(* IEC 61131-3 sources: Test-Git_ESME26/TestProgettoESME_26.fbsproj/PacDriveLib Migration/Motion/Control/PDL_FB_Brake.fb.st^, 4 files *)

(* ---- AsyncExtDiagTranslation.meth.st ---- *)
METHOD AsyncExtDiagTranslation : BOOL
VAR_INPUT
END_VAR

CASE etResult OF
	SE_Async.ET_Result.MaxNumOfReusableObjectsExceeded: ; // No error message. Try again to Start in next cycle

	SE_Async.ET_Result.AsyncAddWasNotSuccessful:
		SetDiagOutput(	i_etDiag	:= GD.ET_Diag.UnexpectedProgramBehavior,
						i_etDiagExt := PDL_ET_DiagExt.AsyncAddWasNotSuccessful,
						i_sMsg		:= SE_CTBX.FC_MultiConcat(	i_sString1 := '#',
														i_sString2 := DINT_TO_STRING(diState),
														i_sString3 := ' G_ifAsync.Start: ',
														i_sString4 := PDL_FC_EtDiagExtToString(etDiagExt)));

	SE_Async.ET_Result.InterfaceCastFailed:
		SetDiagOutput(	i_etDiag	:= GD.ET_Diag.UnexpectedProgramBehavior,
						i_etDiagExt := PDL_ET_DiagExt.InterfaceCastFailed,
						i_sMsg		:= SE_CTBX.FC_MultiConcat(	i_sString1 := '#',
														i_sString2 := DINT_TO_STRING(diState),
														i_sString3 := ' G_ifAsync.Start: ',
														i_sString4 := PDL_FC_EtDiagExtToString(etDiagExt)));

	SE_Async.ET_Result.SemaphoreCreateFailed:
		SetDiagOutput(	i_etDiag	:= GD.ET_Diag.UnexpectedProgramBehavior,
						i_etDiagExt := PDL_ET_DiagExt.SemaphoreMeCreateFailed,
						i_sMsg		:= SE_CTBX.FC_MultiConcat(	i_sString1 := '#',
														i_sString2 := DINT_TO_STRING(diState),
														i_sString3 := ' G_ifAsync.Start: ',
														i_sString4 := PDL_FC_EtDiagExtToString(etDiagExt)));

	SE_Async.ET_Result.AsyncInvalid:
		SetDiagOutput(	i_etDiag	:= GD.ET_Diag.InputParameterInvalid,
						i_etDiagExt := PDL_ET_DiagExt.AsyncInvalid,
						i_sMsg		:= SE_CTBX.FC_MultiConcat(	i_sString1 := '#',
														i_sString2 := DINT_TO_STRING(diState),
														i_sString3 := ' G_ifAsync.Start: ',
														i_sString4 := PDL_FC_EtDiagExtToString(etDiagExt)));

	SE_Async.ET_Result.NoAsyncTasksCreated:
		SetDiagOutput(	i_etDiag	:= GD.ET_Diag.ExecutionAborted,
						i_etDiagExt := PDL_ET_DiagExt.NoAsyncTasksCreated,
						i_sMsg		:= SE_CTBX.FC_MultiConcat(	i_sString1 := '#',
														i_sString2 := DINT_TO_STRING(diState),
														i_sString3 := ' G_ifAsync.Start: ',
														i_sString4 := PDL_FC_EtDiagExtToString(etDiagExt)));

	SE_Async.ET_Result.AsyncInitNotFinished:
		SetDiagOutput(	i_etDiag	:= GD.ET_Diag.ExecutionAborted,
						i_etDiagExt := PDL_ET_DiagExt.AsyncInitNotFinished,
						i_sMsg		:= SE_CTBX.FC_MultiConcat(	i_sString1 := '#',
														i_sString2 := DINT_TO_STRING(diState),
														i_sString3 := ' G_ifAsync.Start: ',
														i_sString4 := PDL_FC_EtDiagExtToString(etDiagExt)));

	SE_Async.ET_Result.ColdResetOfControllerNecessary:
		SetDiagOutput(	i_etDiag	:= GD.ET_Diag.ExecutionAborted,
						i_etDiagExt := PDL_ET_DiagExt.ColdResetOfControllerNecessary,
						i_sMsg		:= SE_CTBX.FC_MultiConcat(	i_sString1 := '#',
														i_sString2 := DINT_TO_STRING(diState),
														i_sString3 := ' G_ifAsync.Start: ',
														i_sString4 := PDL_FC_EtDiagExtToString(etDiagExt)));

	ELSE
		SetDiagOutput(	i_etDiag	:= GD.ET_Diag.UnexpectedProgramBehavior,
						i_etDiagExt := PDL_ET_DiagExt.UnexpectedFeedback,
						i_sMsg		:= SE_CTBX.FC_MultiConcat(	i_sString1 := '#',
														i_sString2 := DINT_TO_STRING(diState),
														i_sString3 := ' G_ifAsync.Start: ',
														i_sString4 := PDL_FC_EtDiagExtToString(etDiagExt)));
END_CASE

(* ---- InitInterfaces.meth.st ---- *)
{attribute 'conditionalshow_all_locals'}
METHOD PRIVATE InitInterfaces : BOOL
VAR_INPUT
END_VAR

InitInterfaces := FALSE;
IF i_ifDrive = 0 THEN
	SetDiagOutput(	i_etDiag	:= GD.ET_Diag.InputParameterInvalid,
					i_etDiagExt := PDL_ET_DiagExt.DriveInvalid,
					i_sMsg		:= 'i_ifDrive - Invalid Interface');
	RETURN;
END_IF

xSuccess := __QUERYINTERFACE(i_ifDrive, ifGetParentDevice);
IF NOT xSuccess OR ifGetParentDevice = 0 THEN
	SetDiagOutput(	i_etDiag	:= GD.ET_Diag.InputParameterInvalid,
					i_etDiagExt := PDL_ET_DiagExt.DriveInvalid,
					i_sMsg		:= 'i_ifDrive - ifGetParentDevice not implemented');
	RETURN;
ELSE
	ifDeviceAccess := ifGetParentDevice.GetParentDevice();
END_IF

xSuccess := __QUERYINTERFACE(ifDeviceAccess,ifBrakeAccess);
IF NOT xSuccess OR ifBrakeAccess = 0 THEN
	SetDiagOutput(	i_etDiag	:= GD.ET_Diag.InputParameterInvalid,
					i_etDiagExt := PDL_ET_DiagExt.DriveInvalid,
					i_sMsg		:= 'i_ifDrive - IF_Brake not implemented');
	RETURN;
END_IF
ifBrake := ifBrakeAccess.Brake;

xSuccess := __QUERYINTERFACE(ifDeviceAccess, ifWorkingModeAccess);
IF NOT xSuccess OR ifWorkingModeAccess = 0 THEN
	SetDiagOutput(	i_etDiag	:= GD.ET_Diag.InputParameterInvalid,
					i_etDiagExt := PDL_ET_DiagExt.DriveInvalid,
					i_sMsg		:= 'i_ifDrive - IF_WorkingMode not implemented');
	RETURN;
END_IF
ifWorkingMode := ifWorkingModeAccess.WorkingMode;

xSuccess := __QUERYINTERFACE(ifDeviceAccess, ifDeviceTreeObjectAccess);
IF xSuccess THEN
	sDriveName := ifDeviceTreeObjectAccess.DeviceTreeObject.Name;
ELSE
	sDriveName := '';
END_IF

InitInterfaces := TRUE;

(* ---- RegisterLoggerPoint.meth.st ---- *)
METHOD PUBLIC RegisterLoggerPoint
VAR_INPUT
	i_ifParent		: APL.IF_LoggerPoint;
	i_sName			: STRING[80];
END_VAR
VAR_OUTPUT
	q_etDiag		: GD.ET_Diag := GD.ET_Diag.Ok;
	q_etDiagExt		: PDL_ET_DiagExt := PDL_ET_DiagExt.Ok;
END_VAR
VAR
	etDiagBuffer		: GD.ET_Diag;
	etDiagExtBufferAPL	: APL.ET_DiagExt;
END_VAR

fbLoggerPoint.RegisterLoggerPoint(	i_ifParent		:= i_ifParent,
									i_sName			:= i_sName,
									i_sType			:= 'FB_Brake',
									i_sSource		:= 'PDL',
									q_etDiag		=> etDiagBuffer,
									q_etDiagExt		=> etDiagExtBufferAPL);
IF (etDiagBuffer <> GD.ET_Diag.Ok) THEN
	CASE etDiagExtBufferAPL OF
		APL.ET_DiagExt.ParentInvalid:
			q_etDiag := GD.ET_Diag.InputParameterInvalid;
			q_etDiagExt := PDL_ET_DiagExt.ParentInvalid;

		APL.ET_DiagExt.ParentNotRegistered:
			q_etDiag := GD.ET_Diag.InputParameterInvalid;
			q_etDiagExt := PDL_ET_DiagExt.ParentNotRegistered;

		APL.ET_DiagExt.MaxNumberOfLoggerPointsExeeded:
			q_etDiag := GD.ET_Diag.InputParameterInvalid;
			q_etDiagExt := PDL_ET_DiagExt.MaxNumberOfLoggerPointsExeeded;

	ELSE
		q_etDiag := GD.ET_Diag.UnexpectedProgramBehavior;
		q_etdiagExt := PDL_ET_DiagExt.UnexpectedDiagExt;
	END_CASE
END_IF

(* ---- SetDiagOutput.meth.st ---- *)
{attribute 'hide'}
METHOD SetDiagOutput : BOOL
VAR_INPUT
	i_etDiag	: GD.ET_Diag;
	i_etDiagExt	: PDL_ET_DiagExt;
	i_sMsg		: STRING[80];
END_VAR
VAR
END_VAR

IF i_etDiag <> GD.ET_Diag.Ok THEN
	q_xReady := FALSE;
END_IF

IF q_etDiag = GD.ET_Diag.OK OR i_etDiagExt = PDL_ET_DiagExt.Disabled THEN

	q_etDiag 	:= i_etDiag;
	q_etDiagExt := i_etDiagExt;
	q_sMsg 		:= i_sMsg;

END_IF
